Staubli VAL3: forItem.pjx

--- forItem.pjx ---
Parameters version=s8.12.1Cs9_BS2449 stackSize=5000 millimeterUnit=true
Data file=forItem.dtx

--- forItem.dtx ---
public num nLoopValue
public bool bIOdisable
public string sIOindex
public string sForTRAJ
